Fanuc KAREL source: kt00069.KL

-- PROVISIONAL review KL for V770-1; original PC SHA256 a2d005a02457169ed1a694cbcf17e393a8d0ce10b1c58b54fc35bb10b154df32
-- Incomplete behavior may be omitted. Consult companion uncertainty JSON. Do not deploy.
PROGRAM KT00069
%NOLOCKGROUP
VAR
  I1 : INTEGER
  OUT : INTEGER
-- UNRESOLVED_DECL Y2 type=002018
BEGIN
  -- UNRESOLVED_PC offsets 5-16; opcodes 2E,23
  -- UNRESOLVED_PC offsets 21-35; opcodes 2E,22,9D,33,B2
  -- UNRESOLVED_PC offsets 40-62; opcodes 21,22,9D,33,B1,54,23
  -- UNRESOLVED_PC offsets 67-71; opcodes 7F
END KT00069
